Staubli VAL3: modifyPara.pgx

public program modifyPara(string x_sKey, num x_nIndex, num x_nMoveType, num x_nParaSpeed, num x_nParaBlend, num x_nParaPercent, string x_sComment, bool x_bSafePoint, string x_sBlend, bool& x_bToSave, num& x_nValue[], num x_nParaAcel)
begin
  trajTemp:tTrajItem[x_sKey].pPointItem[x_nIndex].sID=x_sComment
  trajTemp:tTrajItem[x_sKey].pPointItem[x_nIndex].pParaItem.nMoveType=x_nMoveType
  trajTemp:tTrajItem[x_sKey].pPointItem[x_nIndex].pParaItem.mMdesc.vel=x_nParaSpeed
  trajTemp:tTrajItem[x_sKey].pPointItem[x_nIndex].pParaItem.mMdesc.accel=x_nParaAcel
  trajTemp:tTrajItem[x_sKey].pPointItem[x_nIndex].pParaItem.mMdesc.leave=x_nParaBlend
  trajTemp:tTrajItem[x_sKey].pPointItem[x_nIndex].pParaItem.nPercentage=x_nParaPercent
  trajTemp:tTrajItem[x_sKey].pPointItem.pParaItem.bSafePoint=(x_bSafePoint==true)
  switch x_sBlend
    case "OFF"
      trajTemp:tTrajItem[x_sKey].pPointItem[x_nIndex].pParaItem.mMdesc.blend=off
    break
    case "关节"
      trajTemp:tTrajItem[x_sKey].pPointItem[x_nIndex].pParaItem.mMdesc.blend=joint
    break
    case "笛卡尔"
      trajTemp:tTrajItem[x_sKey].pPointItem[x_nIndex].pParaItem.mMdesc.blend=Cartesian
    break

  endSwitch
  switch x_nMoveType
    case 0
      trajTemp:tTrajItem[x_sKey].pPointItem[x_nIndex].jJointRx.j1=x_nValue[0]
      trajTemp:tTrajItem[x_sKey].pPointItem[x_nIndex].jJointRx.j2=x_nValue[1]
      trajTemp:tTrajItem[x_sKey].pPointItem[x_nIndex].jJointRx.j3=x_nValue[2]
      trajTemp:tTrajItem[x_sKey].pPointItem[x_nIndex].jJointRx.j4=x_nValue[3]
      trajTemp:tTrajItem[x_sKey].pPointItem[x_nIndex].jJointRx.j5=x_nValue[4]
      trajTemp:tTrajItem[x_sKey].pPointItem[x_nIndex].jJointRx.j6=x_nValue[5]
    break
    case 1
      trajTemp:tTrajItem[x_sKey].pPointItem[x_nIndex].pPointRx.trsf.x=x_nValue[0]
      trajTemp:tTrajItem[x_sKey].pPointItem[x_nIndex].pPointRx.trsf.y=x_nValue[1]
      trajTemp:tTrajItem[x_sKey].pPointItem[x_nIndex].pPointRx.trsf.z=x_nValue[2]
      trajTemp:tTrajItem[x_sKey].pPointItem[x_nIndex].pPointRx.trsf.rx=x_nValue[3]
      trajTemp:tTrajItem[x_sKey].pPointItem[x_nIndex].pPointRx.trsf.ry=x_nValue[4]
      trajTemp:tTrajItem[x_sKey].pPointItem[x_nIndex].pPointRx.trsf.rz=x_nValue[5]
    break
    case 2
      trajTemp:tTrajItem[x_sKey].pPointItem[x_nIndex].pPointRx.trsf.x=x_nValue[0]
      trajTemp:tTrajItem[x_sKey].pPointItem[x_nIndex].pPointRx.trsf.y=x_nValue[1]
      trajTemp:tTrajItem[x_sKey].pPointItem[x_nIndex].pPointRx.trsf.z=x_nValue[2]
      trajTemp:tTrajItem[x_sKey].pPointItem[x_nIndex].pPointRx.trsf.rx=x_nValue[3]
      trajTemp:tTrajItem[x_sKey].pPointItem[x_nIndex].pPointRx.trsf.ry=x_nValue[4]
      trajTemp:tTrajItem[x_sKey].pPointItem[x_nIndex].pPointRx.trsf.rz=x_nValue[5]
      trajTemp:tTrajItem[x_sKey].pPointItem[x_nIndex].pInter.trsf.x=x_nValue[6]
      trajTemp:tTrajItem[x_sKey].pPointItem[x_nIndex].pInter.trsf.y=x_nValue[7]
      trajTemp:tTrajItem[x_sKey].pPointItem[x_nIndex].pInter.trsf.z=x_nValue[8]
      trajTemp:tTrajItem[x_sKey].pPointItem[x_nIndex].pInter.trsf.rx=x_nValue[9]
      trajTemp:tTrajItem[x_sKey].pPointItem[x_nIndex].pInter.trsf.ry=x_nValue[10]
      trajTemp:tTrajItem[x_sKey].pPointItem[x_nIndex].pInter.trsf.rz=x_nValue[11]
    break
  endSwitch
  //trajTemp:libSave()
  //delay(0.5)
  logMsg("参数已修改")
  x_bToSave=true
end
